Omron CX-Programmer project  (CX-Programmer ?)

# PLC :  

## Function block LD_Probe
VAR_IN_OUT
  SharedBit : BOOL;
END_VAR

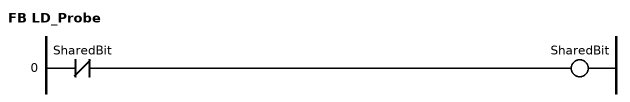
; rung 0
LDNOT SharedBit
OUT SharedBit